Yaskawa INFORM job: 1-DEFRO-60.JBI

/JOB
//NAME 1-DEFRO-60
//POS
///NPOS 0,0,0,0,0,0
//INST
///DATE 2025/01/10 11:18
///ATTR SC,RW,CJ
///GROUP1 RB1,BS1,ST3
NOP
END
